    M_PRO_CHARGING_SYSTEMS_1623 : UINT := 1623; (* Manufacturer: PRO Charging Systems, LLC | Location: La Vergne, TN, USA - 2026-01-27 *)
    M_CROSSCONTROL : UINT := 1624; (* Manufacturer: CrossControl | Location: Alfta, Sweden - 2026-01-27 *)
    M_DMX_POWER : UINT := 1625; (* Manufacturer: DMX Power LLC | Location: Oakdale, MN, USA - 2026-01-27 *)
    M_SMP_STABIL : UINT := 1626; (* Manufacturer: SMP STABIL GmbH | Location: Pécel, Hungary - 2026-01-27 *)
    M_ROTER_ITALIA : UINT := 1627; (* Manufacturer: Roter Italia | Location: Ostiglia(MN), Italy - 2026-01-27 *)
    M_VANEMAR : UINT := 1628; (* Manufacturer: Vanemar, Inc. | Location: Fort Lauderdale, FL, USA - 2026-01-27 *)
    M_DSPACE_SE_AND : UINT := 1629; (* Manufacturer: dSPACE SE & Co. KG | Location: Paderborn, North Rhine Westphalia, Germany - *)
    M_RAINER_MEYER_LANDMASCHINEN : UINT := 1630; (* Manufacturer: Rainer Meyer Landmaschinen GmbH | Location: Niedersachsen, Germany - 2026-01-27 *)
    M_LEIDOS : UINT := 1631; (* Manufacturer: Leidos | Location: Reston, VA, USA - 2026-01-27 *)
    M_ZOCON : UINT := 1632; (* Manufacturer: Zocon | Location: Joure, The Netherlands - 2026-02-09 *)
    M_ZYDRO_MARINE_TECHNOLOGIES : UINT := 1633; (* Manufacturer: Zydro Marine Technologies, Inc. | Location: Boston, MA, USA - 2026-02-09 *)
    M_IBISUL_ELETR_NICA_LTDA : UINT := 1634; (* Manufacturer: IBISUL ELETRÔNICA LTDA | Location: Ibirubá, Rio Grande do Sul, Brazil - 2026-02-09 *)
    M_SAFRAMAX_INDUSTRIAL : UINT := 1635; (* Manufacturer: Saframax Industrial | Location: Campo Mourão, Paraná, Brazil - 2026-02-09 *)
    M_TBB_POWER : UINT := 1636; (* Manufacturer: TBB POWER (XIAMEN) Co., Ltd. | Location: Xiamen, Fujian, China - 2026-02-13 *)
    M_SCHERZINGER_PUMPEN_AND : UINT := 1637; (* Manufacturer: Scherzinger Pumpen GmbH & Co. KG | Location: Furtwangen im Schwarzwald, *)
    M_TEMPA_TEKNIK : UINT := 1638; (* Manufacturer: TEMPA TEKNIK | Location: Tekirdag, Turkey - 2026-02-18 *)
    M_GEA_FARM_TECHNOLOGIES_CANADA : UINT := 1639; (* Manufacturer: GEA Farm Technologies Canada Inc. | Location: Drummondville, QC, Canada - *)
    M_PEIKA : UINT := 1640; (* Manufacturer: PEIKA | Location: Bydgoszcz, Kujawsko-Pomorskie, Poland - 2026-04-02 *)
    M_LITHOS_ENERGY : UINT := 1641; (* Manufacturer: Lithos Energy | Location: Hayward, CA, USA - 2026-04-02 *)
    M_KW_GENERATOR : UINT := 1642; (* Manufacturer: KW-Generator GmbH | Location: Schwäbisch Gmünd, Baden-Württemberg, Germany *)
    M_CRMR_TECHNOLOGY : UINT := 1643; (* Manufacturer: CRMR Technology, Inc. | Location: Miami, FL, USA - 2026-04-02 *)
    M_U_AND_R_GMBH_HARDWARE_UND_SYSTEMDESIGN : UINT := 1644; (* Manufacturer: U&R GmbH Hardware- und Systemdesign | Location: Erbach, Baden-Wuerttemberg *)
    M_DC_ELECTRONICS : UINT := 1645; (* Manufacturer: DC Electronics | Location: Maldon, Essex, UK - 2026-04-02 *)
    M_WATT_AND_SEA : UINT := 1646; (* Manufacturer: WATT AND SEA | Location: La Rochelle, France - 2026-04-02 *)
    M_NOVATRON_OY : UINT := 1647; (* Manufacturer: Novatron Oy | Location: Pirkkala, Pirkanmaa, Finland - 2026-04-02 *)
    M_ALTEK : UINT := 1648; (* Manufacturer: Altek GmbH | Location: Rottenburg, BW, Germany - 2026-07-23 *)
    M_STARTER_AND_GENERATOR_EXCHANGE_SERVICE : UINT := 1649; (* Manufacturer: Starter & Generator Exchange Service Pty Ltd | Location: Brisbane, Queensland *)
    M_SHANGHAI_INFIPAX_TECHNOLOGY : UINT := 1650; (* Manufacturer: Shanghai Infipax Technology Co., Ltd. | Location: Shanghai, China - 2026-07-23 *)
    M_CREATIVE_WERKS : UINT := 1651; (* Manufacturer: Creative Werks Inc. | Location: Des Moines, IA, USA - 2026-04-02 *)
    M_COSTRUZIONI_MOTORI_DIESEL : UINT := 1652; (* Manufacturer: Costruzioni Motori Diesel (CMD) | Location: San Nicola La Strada, CA, Italy *)
    M_SCHAFFER_FARMING_TECHNOLOGIES : UINT := 1653; (* Manufacturer: Schaffer Farming Technologies | Location: Mercer, PA, USA - 2026-04-02 *)
    M_INVENTURE_ELECTRONICS : UINT := 1654; (* Manufacturer: Inventure Electronics | Location: Goshen, IN, USA - 2026-05-06 *)
    M_ELECTROSEA : UINT := 1655; (* Manufacturer: Electrosea | Location: Plymouth, MN, USA - 2026-05-06 *)
    M_SUPERSTREAM_OY : UINT := 1656; (* Manufacturer: Superstream Oy | Location: Helsinki, Finland - 2026-07-23 *)
    M_ISRINGHAUSEN_GMBH_AND : UINT := 1657; (* Manufacturer: ISRINGHAUSEN GmbH & Co. KG | Location: Lemgo, Germany - 2026-05-06 *)
    M_ROUSH : UINT := 1658; (* Manufacturer: Roush | Location: Livonia, MI, USA - 2026-05-06 *)
    M_TSM_SENSORS_S_R_L : UINT := 1659; (* Manufacturer: TSM Sensors S.r.l. | Location: Erbusco, Italy - 2026-05-06 *)
    M_ARETE_KLEJBUK_SPOLKA_JAWNA : UINT := 1660; (* Manufacturer: ARETE Klejbuk Spolka Jawna | Location: Choroszcz, Poland - 2026-05-06 *)
    M_CEFIROS : UINT := 1661; (* Manufacturer: CEFIROS | Location: Cordoba, Argentina - 2026-05-06 *)
    M_REMOTE_CONTROL_TECHNOLOGIES : UINT := 1662; (* Manufacturer: Remote Control Technologies (RCT) | Location: Perth, WA, Australia - 2026-05-06 *)
    M_WANDFLUH_AG : UINT := 1663; (* Manufacturer: Wandfluh AG | Location: Frutigen, BE, Switzerland - 2026-05-12 *)
    M_NAUTECH : UINT := 1664; (* Manufacturer: Nautech Ltd. | Location: Balatonfured, Hungary - 2026-07-23 *)
    M_ICP_SYSTEMS_B_V : UINT := 1665; (* Manufacturer: ICP Systems B.V. | Location: Holten, Overijssel, Netherlands - 2026-07-23 *)
    M_TERSUS_GNSS : UINT := 1666; (* Manufacturer: Tersus GNSS Inc. | Location: Shanghai, China - 2026-07-23 *)
    M_ADVANCED_FLOW_SOLUTIONS : UINT := 1667; (* Manufacturer: Advanced Flow Solutions, Inc. | Location: Oklahoma City, OK, USA - 2026-07-23 *)
    M_PERFECT_PRECISION_AGRICULTURE : UINT := 1668; (* Manufacturer: Perfect Precision Agriculture | Location: Dundee, KZN, South Africa - 2026-08-04 *)
    M_SHENZHEN_TOPBAND : UINT := 1669; (* Manufacturer: Shenzhen Topband Co. Ltd. | Location: Shiyan, Guangdong Province, China *)
    M_MCT_TECHNIC_SENSOR_A_S : UINT := 1670; (* Manufacturer: MCT TECHNIC SENSOR A.S. | Location: Bakirkoy, Istanbul, Turkey - 2026-07-23 *)
    M_LOOKOUT : UINT := 1671; (* Manufacturer: LOOKOUT | Location: Somerville, MA, USA - 2026-07-23 *)
    M_ANDREAS_LUPOLD_HYDROTECHNIK : UINT := 1672; (* Manufacturer: Andreas Lupold Hydrotechnik GmbH | Location: Voehringen, BW, Germany - 2026-07-23 *)
    M_SISTEMATICA_S_R_L : UINT := 1673; (* Manufacturer: SISTEMATICA S.r.l | Location: Turin, Italy - 2026-07-23 *)
    M_YACHTWAVE : UINT := 1674; (* Manufacturer: YACHTWAVE | Location: Sarasota, FL, USA - 2026-07-23 *)
    M_TETRADYNE : UINT := 1675; (* Manufacturer: Tetradyne Co., Ltd. | Location: Seoul, South Korea - 2026-07-23 *)
    M_MERLIN_SOLAR_TECHNOLOGIES : UINT := 1676; (* Manufacturer: Merlin Solar Technologies, Inc. | Location: San Jose, California, USA *)
    M_GINT : UINT := 1684; (* Manufacturer: GINT Co., Ltd. | Location: Seongnam-si, Gyeonggi-do, Republic of Korea *)
    M_TANIE_NAWIGOWANIE : UINT := 1685; (* Manufacturer: Tanie Nawigowanie | Location: Wroclaw, Poland - 2026-09-24 *)
    M_PTM_S_R_L : UINT := 1695; (* Manufacturer: PTM S.r.l. | Location: Visano, Italy - 2026-09-24 *)
    M_COMESYS : UINT := 1700; (* Manufacturer: ComeSys Ltd. | Location: Busan, South Korea - 2026-11-12 *)
    M_INNOV_GPS : UINT := 1704; (* Manufacturer: INNOV.GPS | Location: Villers les Cagnicourt, France - 2026-11-12 *)
    M_OPTISENS_INTELLIGENT_TECHNOLOGY : UINT := 1712; (* Manufacturer: Optisens Intelligent Technology Co., Ltd. | Location: Shanghai, China *)
    M_SEASTAR_SOLUTIONS : UINT := 1850; (* Manufacturer: Seastar Solutions (formerly Teleflex) | Location: Litchfield, IL - 2021-08-26 *)
    M_RAYMARINE : UINT := 1851; (* Manufacturer: RayMarine | Location: Portsmouth, Hampshire UK - 2003-07-20 *)
    M_NAVIONICS : UINT := 1852; (* Manufacturer: Navionics | Location: Wareham, MA USA - 2003-07-20 *)
    M_JAPAN_RADIO : UINT := 1853; (* Manufacturer: Japan Radio Co | Location: Seattle, WA USA - 2003-07-20 *)
    M_NORTHSTAR_TECHNOLOGIES : UINT := 1854; (* Manufacturer: Northstar Technologies | Location: Acton, MA USA - 2003-07-20 *)
    M_FURUNO_USA : UINT := 1855; (* Manufacturer: Furuno USA | Location: Camas, WA USA - 2003-07-20 *)
    M_TRIMBLE : UINT := 1856; (* Manufacturer: Trimble | Location: Sunnyvale, CA USA - 2003-07-20 *)
    M_SIMRAD : UINT := 1857; (* Manufacturer: Simrad | Location: Egersund, Norway - 2003-07-20 *)
    M_LITTON : UINT := 1858; (* Manufacturer: Litton | Location: Charlottesville, VA USA - 2003-07-20 *)
    M_KVASAR : UINT := 1859; (* Manufacturer: Kvasar AB | Location: Kinnahult, Sweden - 2003-07-20 *)
    M_MMP : UINT := 1860; (* Manufacturer: MMP | Location: Fircrest, WA USA - 2003-07-20 *)
    M_VECTOR_NORTH_AMERICA : UINT := 1861; (* Manufacturer: Vector North America (formerly Vector Cantech) | Location: Novi, MI USA - *)
    M_SANSHIN : UINT := 1862; (* Manufacturer: Sanshin | Location: Shizuoka, Japan - 2003-07-20 *)
    M_THOMAS_G_FARIA : UINT := 1863; (* Manufacturer: Thomas G. Faria Co. | Location: Uncasville, CT USA - 2003-07-20 *)
  END_VAR
END_GLOBALCONSTANTS
